INTERFACE I_SpeedController

METHOD PUBLIC JogFwd
END_METHOD

METHOD PUBLIC JogRev
END_METHOD

METHOD PUBLIC LatchJogFwd
END_METHOD

METHOD PUBLIC LatchJogRev
END_METHOD

METHOD PUBLIC ReadStatus : ST_SpeedControllerStatus
END_METHOD

METHOD PUBLIC Reset
END_METHOD

METHOD PUBLIC SetMotionParam 
VAR_INPUT
	param		: E_MotorMotionParam;
	val			: LREAL;
END_VAR
END_METHOD

METHOD PUBLIC Stop
END_METHOD

END_INTERFACE

(* stored: Version 1.1.0.1, ProductVersion 3.1.4024.12
   Itf I_SpeedController: Id {bf7b357c-8a33-46d9-bc9a-ccb99e6b4603}
   Method JogFwd: Id {296c72fb-1c8b-4f55-91b2-1658ca46a4fd}
   Method JogRev: Id {8bb0f188-78f8-43df-8726-8dc8a4ad7ba2}
   Method LatchJogFwd: Id {77c4995b-fa10-4390-b33f-c60fc71adffc}
   Method LatchJogRev: Id {5c3129c1-35ee-473e-a8b0-9aae7c77e60e}
   Method ReadStatus: Id {5e803f8f-4d8d-438e-a37d-0263051e497c}
   Method Reset: Id {f8d4cc7c-5608-4a57-88af-4e178509b3fa}
   Method SetMotionParam: Id {a6fcd93d-5411-4c81-8649-16d5a2f69728}
   Method Stop: Id {c66cd3c2-1771-4893-bc77-08dc38c112dd} *)
